Fanuc KAREL source: kd00002.KL

PROGRAM KD00002
%STACKSIZE=65535
%PRIORITY=65535
%NOLOCKGROUP
VAR
I : INTEGER
J : INTEGER
B : BOOLEAN
R : REAL
S : STRING[80]
BEGIN
I=1
END KD00002
